{attribute 'TcGvlVarFlags' := 'OPC'}
VAR_GLOBAL
    // Commands — written by Python over ADS, sent to device every cycle
    // ADS symbol: GVL_MenteeMotor.stCmd
    stCmd               : ST_MenteeMotorCmd;

    // Status — read from device every cycle, read by Python over ADS
    // ADS symbol: GVL_MenteeMotor.stStatus
    stStatus            : ST_MenteeMotorStatus;
END_VAR

(* stored: Version 1.1.0.1, ProductVersion 3.1.4026.18
   GVL GVL_MenteeMotor: Id {6c48deb4-c334-4be6-b5b1-49fe7ed0ee96} *)
